PROGRAM POU
VAR
	fOneFloat : REAL;
	sThisIsAString : STRING;
	nAnInteger : INT;
	
	nReturnedNumberOfBytesForFloat : UDINT;
	nReturnedNumberOfBytesForString : UDINT;
	nReturnedNumberOfBytesForInteger : UDINT;
END_VAR

nReturnedNumberOfBytesForFloat := SIZEOF(fOneFloat);
nReturnedNumberOfBytesForString := SIZEOF(sThisIsAString);
nReturnedNumberOfBytesForInteger := SIZEOF(nAnInteger);

END_PROGRAM

(* stored: Version 1.1.0.1
   POU POU: Id {80087357-1119-4c5b-b325-82337c9a2f5c}, SpecialFunc None *)
